Fanuc KAREL source: kb00031.KL

-- PROVISIONAL review KL for V770-1; original PC SHA256 bcb9109cd55f963f44bca0e04bfedaedf411f71fed9a110c99cf2bb49d1f7c0c
-- Incomplete behavior may be omitted. Consult companion uncertainty JSON. Do not deploy.
PROGRAM KB00031
%NOLOCKGROUP
BEGIN
  -- UNRESOLVED_PC offsets 5-16; opcodes 2E,23
  -- UNRESOLVED_PC offsets 21-30; opcodes 3F,75
  -- UNRESOLVED_PC offsets 35-42; opcodes 9D,23
  -- UNRESOLVED_PC offsets 47-71; opcodes 27,22,22,2A,22,31
  -- UNRESOLVED_PC offsets 76-80; opcodes 7F
END KB00031
